FUNCTION_BLOCK DivDez2 (* Dois valores INT em decimos para REAL (/10) *)
  (* Standard: 61499-2 *)
  (* Version 1.0, 04/11/2026, Hidryco, Hidryco, 1.0: OUT1 = IN1 / 10, OUT2 = IN2 / 10. No FieldSignals: corrente (0,1 A) e rotacao (0,1 Hz) dos sopradores Sulzer. *)
  PACKAGE SE.Nereda;
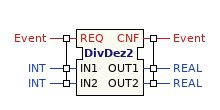
  EVENT_INPUT
    REQ WITH IN1, IN2; (* Converte *)
  END_EVENT
  EVENT_OUTPUT
    CNF WITH OUT1, OUT2; (* Valores convertidos *)
  END_EVENT
  VAR_INPUT
    IN1 : INT; (* Valor em decimos *)
    IN2 : INT; (* Valor em decimos *)
  END_VAR
  VAR_OUTPUT
    OUT1 : REAL; (* IN1 / 10 *)
    OUT2 : REAL; (* IN2 / 10 *)
  END_VAR
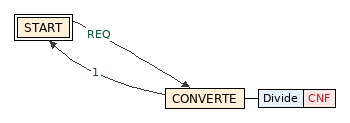
  EC_STATES
    START; (* Estado inicial *)
    CONVERTE : Divide -> CNF; (* Divide por 10 *)
  END_STATES
  EC_TRANSITIONS
    START TO CONVERTE := REQ;
    CONVERTE TO START := 1;
  END_TRANSITIONS
  ALGORITHM Divide IN ST: (* Decimos para unidade *)
OUT1 := INT_TO_REAL(IN1) / 10.0;
OUT2 := INT_TO_REAL(IN2) / 10.0;
  END_ALGORITHM
END_FUNCTION_BLOCK
